(* IEC 61131-3 sources: PLC-Static-Analysis/modules/plc-rules/src/test/resources/PLCA-P006, 2 files *)

(* ---- compliant.st ---- *)
PROGRAM P_NoJump
VAR
    nStep : INT;
END_VAR
IF nStep <> 0 THEN
    nStep := nStep + 1;
END_IF
END_PROGRAM

(* ---- noncompliant.st ---- *)
PROGRAM P_Jump
VAR
    nStep : INT;
END_VAR
IF nStep = 0 THEN
    JMP lEnd; // PLCA-P006
END_IF
nStep := nStep + 1;
lEnd:
END_PROGRAM
